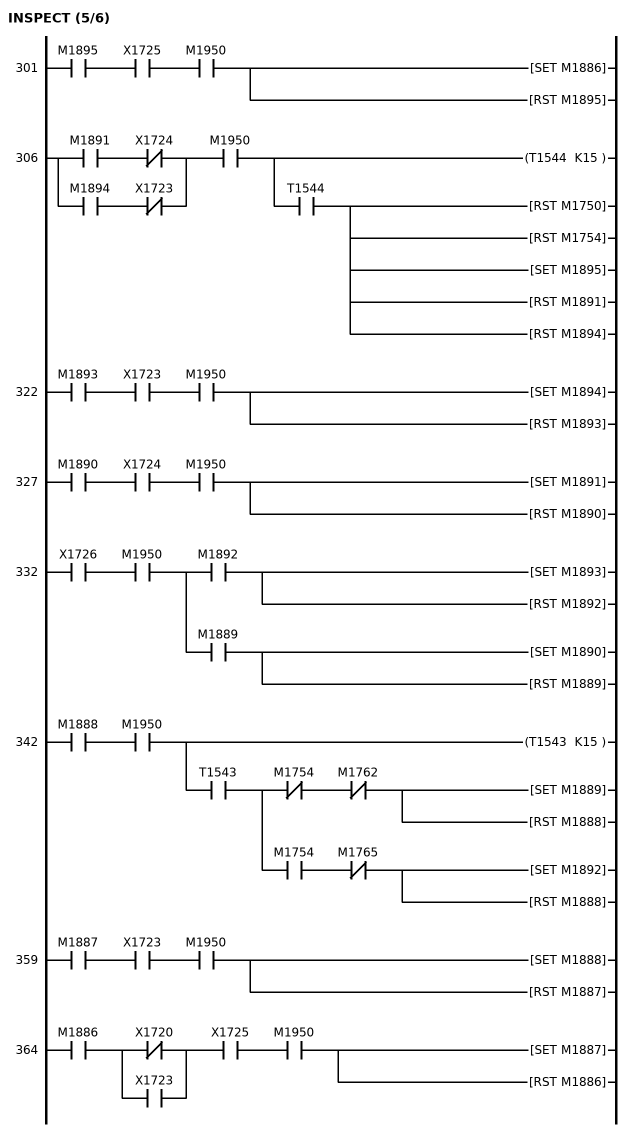
[picture p24: ladder of INSPECT, rungs at steps 301 to 364]
301   LD      M1895
      AND     X1725
      AND     M1950
      SET     M1886
      RST     M1895
306   LD      M1891
      ANI     X1724
      LD      M1894
      ANI     X1723
      ORB
      AND     M1950
      OUT     T1544 K15
      AND     T1544
      RST     M1750
      RST     M1754
      SET     M1895
      RST     M1891
      RST     M1894
322   LD      M1893
      AND     X1723
      AND     M1950
      SET     M1894
      RST     M1893
327   LD      M1890
      AND     X1724
      AND     M1950
      SET     M1891
      RST     M1890
332   LD      X1726
      AND     M1950
      MPS
      AND     M1892
      SET     M1893
      RST     M1892
      MPP
      AND     M1889
      SET     M1890
      RST     M1889
342   LD      M1888
      AND     M1950
      OUT     T1543 K15
      AND     T1543
      MPS
      ANI     M1754
      ANI     M1762
      SET     M1889
      RST     M1888
      MPP
      AND     M1754
      ANI     M1765
      SET     M1892
      RST     M1888
359   LD      M1887
      AND     X1723
      AND     M1950
      SET     M1888
      RST     M1887
364   LD      M1886
      LDI     X1720
      OR      X1723
      ANB
      AND     X1725
      AND     M1950
      SET     M1887
      RST     M1886
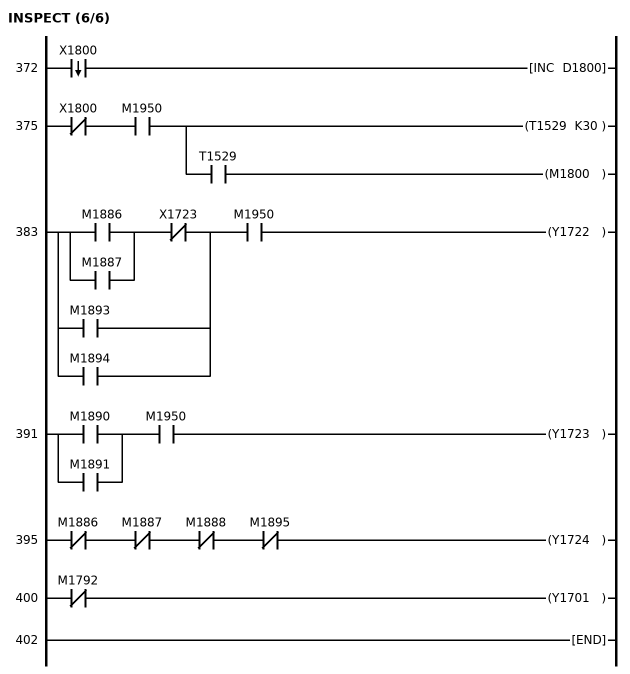
372   LDF     X1800
      INC     D1800
375   LDI     X1800
      AND     M1950
      OUT     T1529 K30
      AND     T1529
      OUT     M1800
383   LD      M1886
      OR      M1887
      ANI     X1723
      LD      M1893
      OR      M1894
      ORB
      AND     M1950
      OUT     Y1722
391   LD      M1890
      OR      M1891
      AND     M1950
      OUT     Y1723
395   LDI     M1886
      ANI     M1887
      ANI     M1888
      ANI     M1895
      OUT     Y1724
400   LDI     M1792
      OUT     Y1701
402   END
END_PROGRAM

PROGRAM RETEST
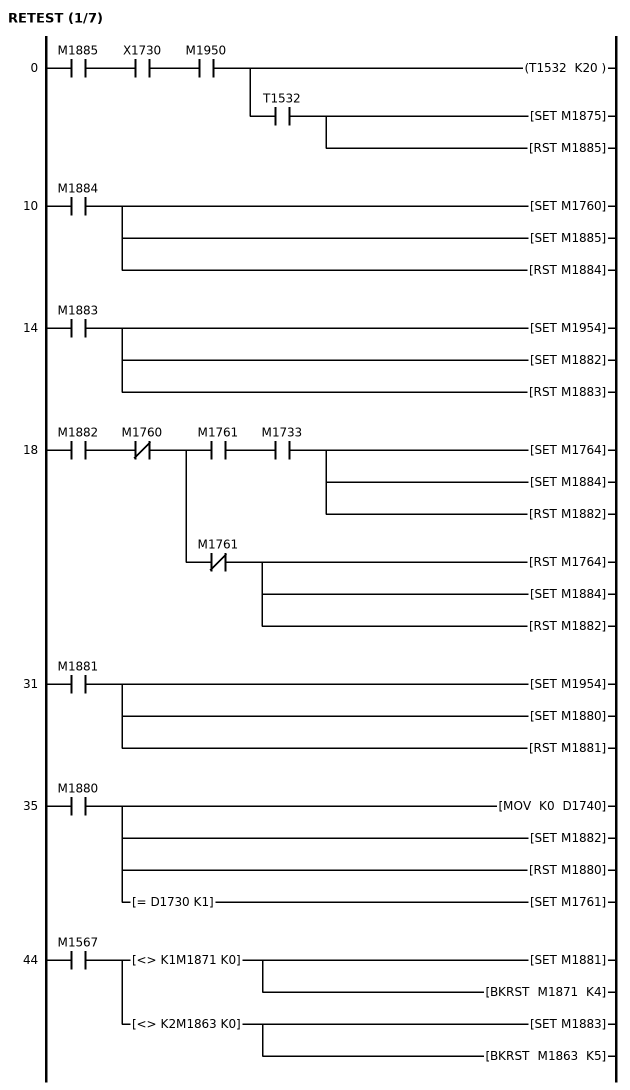
0     LD      M1885
      AND     X1730
      AND     M1950
      OUT     T1532 K20
      AND     T1532
      SET     M1875
      RST     M1885
10    LD      M1884
      SET     M1760
      SET     M1885
      RST     M1884
14    LD      M1883
      SET     M1954
      SET     M1882
      RST     M1883
18    LD      M1882
      ANI     M1760
      MPS
      AND     M1761
      AND     M1733
      SET     M1764
      SET     M1884
      RST     M1882
      MPP
      ANI     M1761
      RST     M1764
      SET     M1884
      RST     M1882
31    LD      M1881
      SET     M1954
      SET     M1880
      RST     M1881
35    LD      M1880
      MOV     K0 D1740
      SET     M1882
      RST     M1880
      AND=    D1730 K1
      SET     M1761
44    LD      M1567
      MPS
      AND<>   K1M1871 K0
      SET     M1881
      BKRST   M1871 K4
      MPP
      AND<>   K2M1863 K0
      SET     M1883
      BKRST   M1863 K5
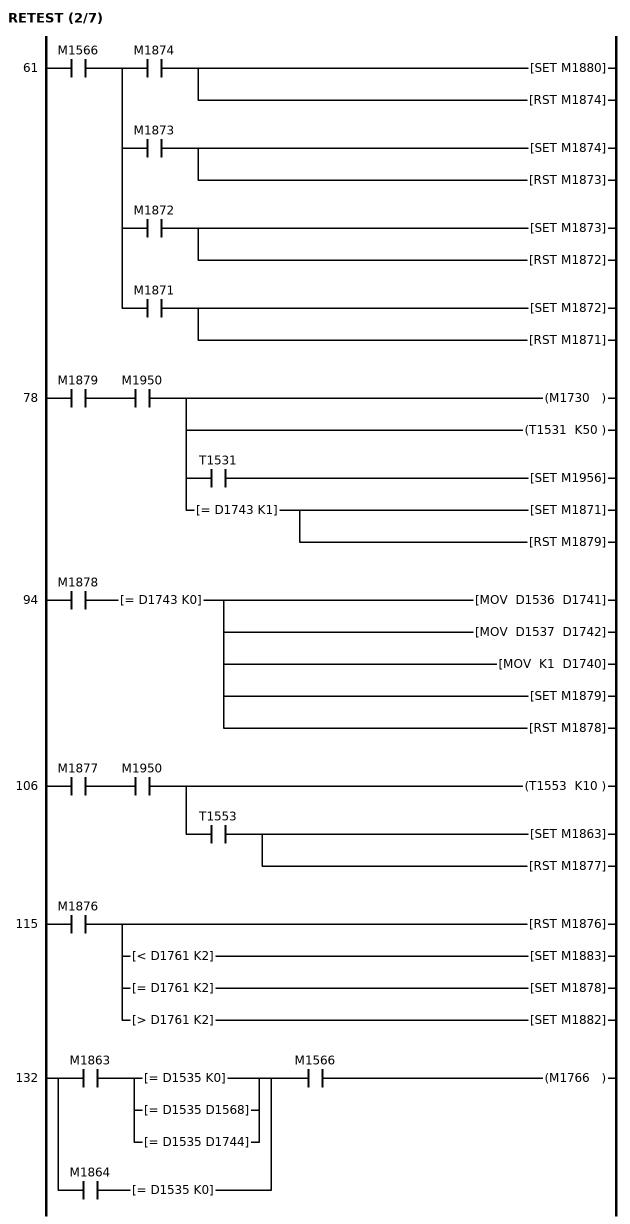
61    LD      M1566
      MPS
      AND     M1874
      SET     M1880
      RST     M1874
      MRD
      AND     M1873
      SET     M1874
      RST     M1873
      MRD
      AND     M1872
      SET     M1873
      RST     M1872
      MPP
      AND     M1871
      SET     M1872
      RST     M1871
78    LD      M1879
      AND     M1950
      OUT     M1730
      OUT     T1531 K50
      MPS
      AND     T1531
      SET     M1956
      MPP
      AND=    D1743 K1
      SET     M1871
      RST     M1879
94    LD      M1878
      AND=    D1743 K0
      MOV     D1536 D1741
      MOV     D1537 D1742
      MOV     K1 D1740
      SET     M1879
      RST     M1878
106   LD      M1877
      AND     M1950
      OUT     T1553 K10
      AND     T1553
      SET     M1863
      RST     M1877
115   LD      M1876
      RST     M1876
      MPS
      AND<    D1761 K2
      SET     M1883
      MRD
      AND=    D1761 K2
      SET     M1878
      MPP
      AND>    D1761 K2
      SET     M1882
132   LD      M1863
      LD=     D1535 K0
      OR=     D1535 D1568
      OR=     D1535 D1744
      ANB
      LD      M1864
      AND=    D1535 K0
      ORB
      AND     M1566
      OUT     M1766
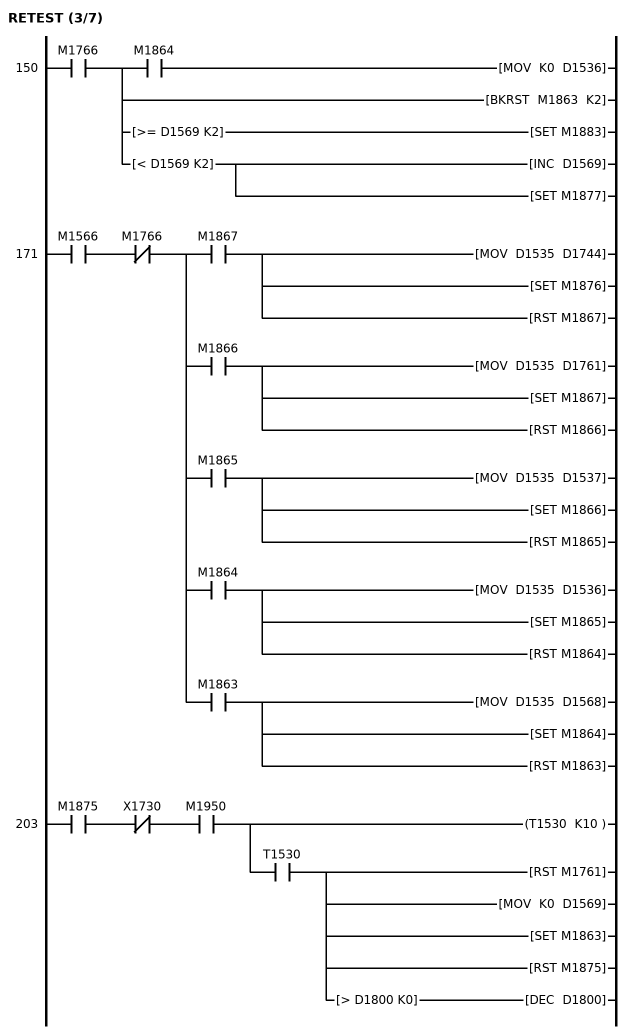
150   LD      M1766
      MPS
      AND     M1864
      MOV     K0 D1536
      MPP
      BKRST   M1863 K2
      MPS
      AND>=   D1569 K2
      SET     M1883
      MPP
      AND<    D1569 K2
      INC     D1569
      SET     M1877
171   LD      M1566
      ANI     M1766
      MPS
      AND     M1867
      MOV     D1535 D1744
      SET     M1876
      RST     M1867
      MRD
      AND     M1866
      MOV     D1535 D1761
      SET     M1867
      RST     M1866
      MRD
      AND     M1865
      MOV     D1535 D1537
      SET     M1866
      RST     M1865
      MRD
      AND     M1864
      MOV     D1535 D1536
      SET     M1865
      RST     M1864
      MPP
      AND     M1863
      MOV     D1535 D1568
      SET     M1864
      RST     M1863
203   LD      M1875
      ANI     X1730
      AND     M1950
      OUT     T1530 K10
      AND     T1530
      RST     M1761
      MOV     K0 D1569
      SET     M1863
      RST     M1875
      AND>    D1800 K0
      DEC     D1800
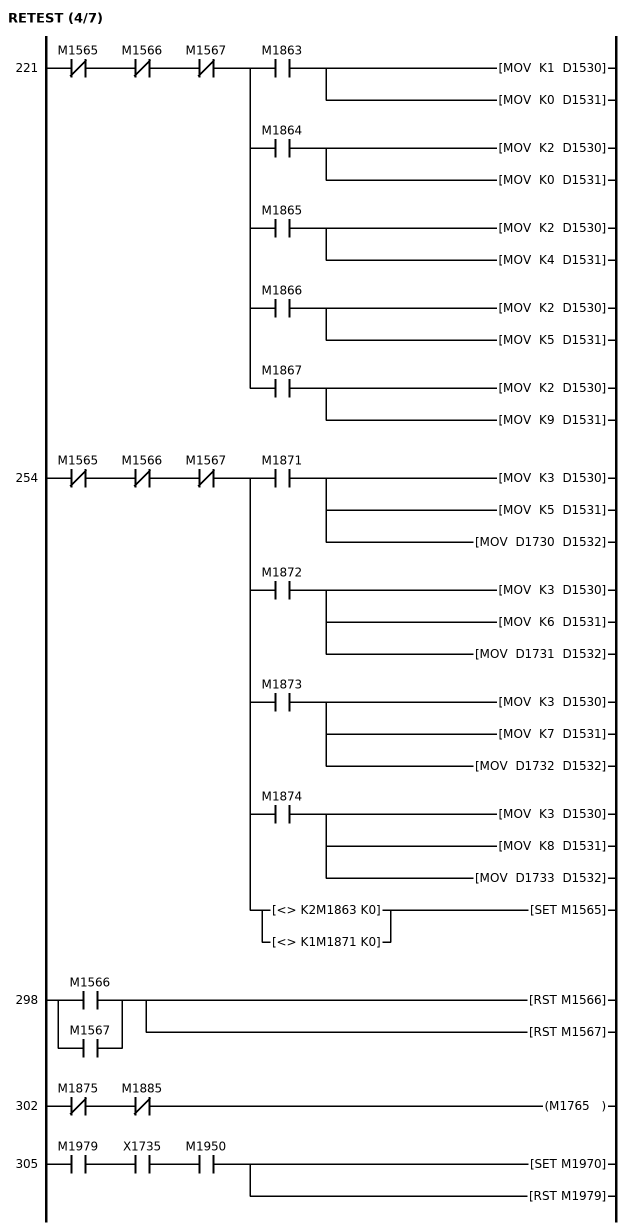
221   LDI     M1565
      ANI     M1566
      ANI     M1567
      MPS
      AND     M1863
      MOV     K1 D1530
      MOV     K0 D1531
      MRD
      AND     M1864
      MOV     K2 D1530
      MOV     K0 D1531
      MRD
      AND     M1865
      MOV     K2 D1530
      MOV     K4 D1531
      MRD
      AND     M1866
      MOV     K2 D1530
      MOV     K5 D1531
      MPP
      AND     M1867
      MOV     K2 D1530
      MOV     K9 D1531
254   LDI     M1565
      ANI     M1566
      ANI     M1567
      MPS
      AND     M1871
      MOV     K3 D1530
      MOV     K5 D1531
      MOV     D1730 D1532
      MRD
      AND     M1872
      MOV     K3 D1530
      MOV     K6 D1531
      MOV     D1731 D1532
      MRD
      AND     M1873
      MOV     K3 D1530
      MOV     K7 D1531
      MOV     D1732 D1532
      MRD
      AND     M1874
      MOV     K3 D1530
      MOV     K8 D1531
      MOV     D1733 D1532
      MPP
      LD<>    K2M1863 K0
      OR<>    K1M1871 K0
      ANB
      SET     M1565
298   LD      M1566
      OR      M1567
      RST     M1566
      RST     M1567
302   LDI     M1875
      ANI     M1885
      OUT     M1765
305   LD      M1979
      AND     X1735
      AND     M1950
      SET     M1970
      RST     M1979
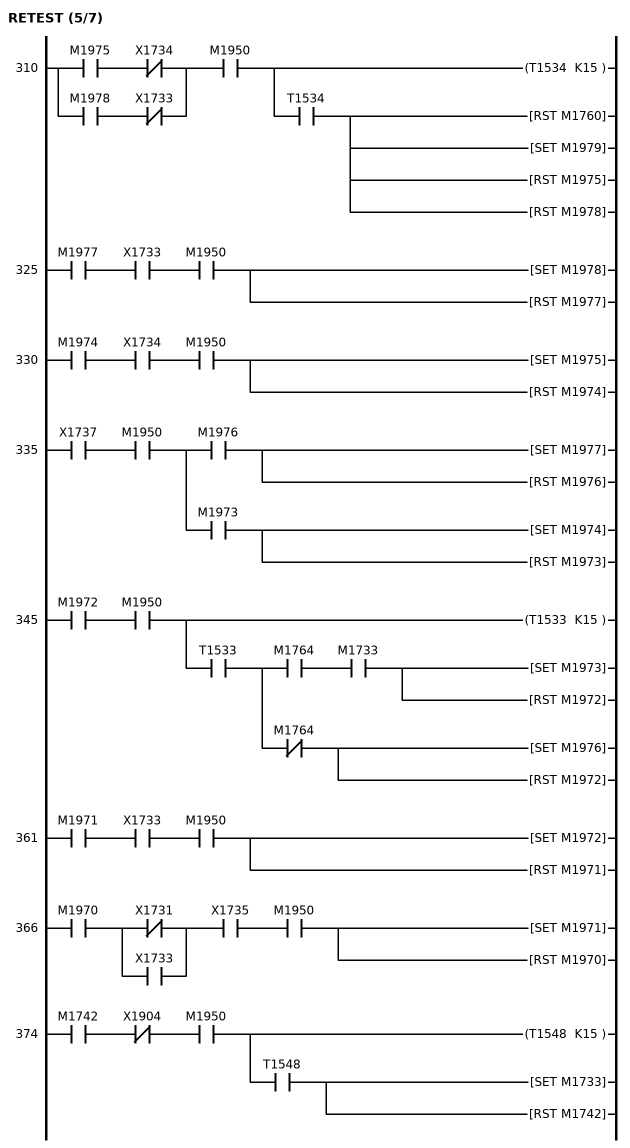
310   LD      M1975
      ANI     X1734
      LD      M1978
      ANI     X1733
      ORB
      AND     M1950
      OUT     T1534 K15
      AND     T1534
      RST     M1760
      SET     M1979
      RST     M1975
      RST     M1978
325   LD      M1977
      AND     X1733
      AND     M1950
      SET     M1978
      RST     M1977
330   LD      M1974
      AND     X1734
      AND     M1950
      SET     M1975
      RST     M1974
335   LD      X1737
      AND     M1950
      MPS
      AND     M1976
      SET     M1977
      RST     M1976
      MPP
      AND     M1973
      SET     M1974
      RST     M1973
345   LD      M1972
      AND     M1950
      OUT     T1533 K15
      AND     T1533
      MPS
      AND     M1764
      AND     M1733
      SET     M1973
      RST     M1972
      MPP
      ANI     M1764
      SET     M1976
      RST     M1972
361   LD      M1971
      AND     X1733
      AND     M1950
      SET     M1972
      RST     M1971
366   LD      M1970
      LDI     X1731
      OR      X1733
      ANB
      AND     X1735
      AND     M1950
      SET     M1971
      RST     M1970
374   LD      M1742
      ANI     X1904
      AND     M1950
      OUT     T1548 K15
      AND     T1548
      SET     M1733
      RST     M1742
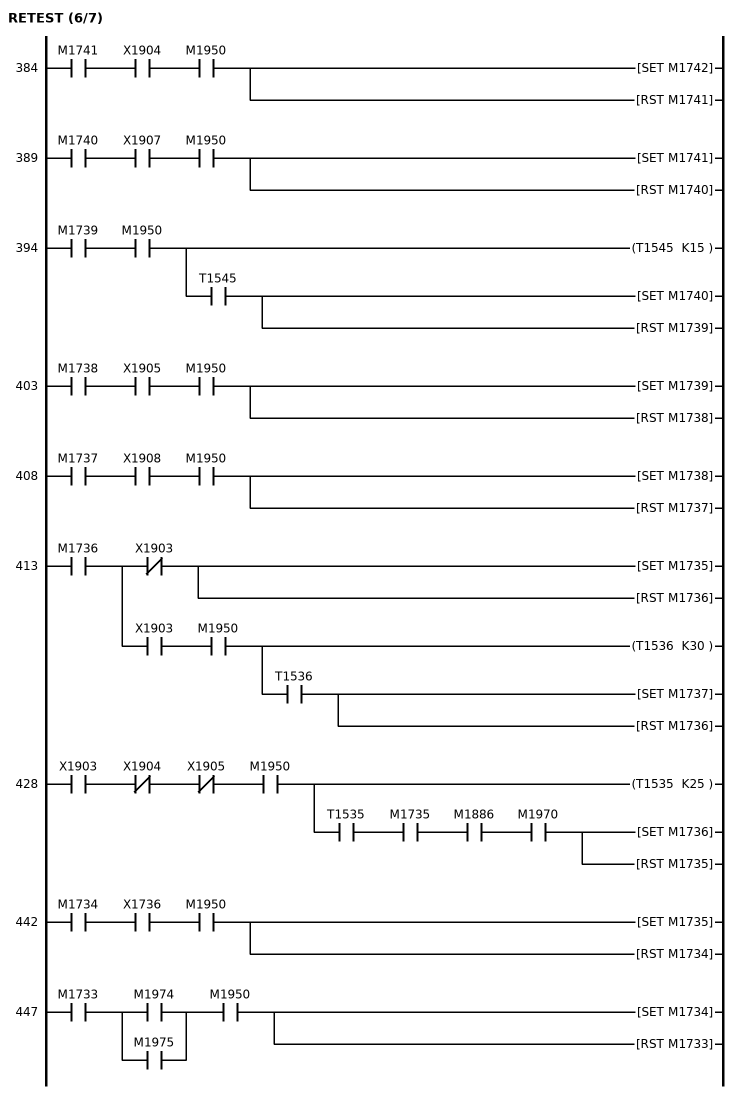
384   LD      M1741
      AND     X1904
      AND     M1950
      SET     M1742
      RST     M1741
389   LD      M1740
      AND     X1907
      AND     M1950
      SET     M1741
      RST     M1740
394   LD      M1739
      AND     M1950
      OUT     T1545 K15
      AND     T1545
      SET     M1740
      RST     M1739
403   LD      M1738
      AND     X1905
      AND     M1950
      SET     M1739
      RST     M1738
408   LD      M1737
      AND     X1908
      AND     M1950
      SET     M1738
      RST     M1737
413   LD      M1736
      MPS
      ANI     X1903
      SET     M1735
      RST     M1736
      MPP
      AND     X1903
      AND     M1950
      OUT     T1536 K30
      AND     T1536
      SET     M1737
      RST     M1736
428   LD      X1903
      ANI     X1904
      ANI     X1905
      AND     M1950
      OUT     T1535 K25
      AND     T1535
      AND     M1735
      AND     M1886
      AND     M1970
      SET     M1736
      RST     M1735
442   LD      M1734
      AND     X1736
      AND     M1950
      SET     M1735
      RST     M1734
447   LD      M1733
      LD      M1974
      OR      M1975
      ANB
      AND     M1950
      SET     M1734
      RST     M1733
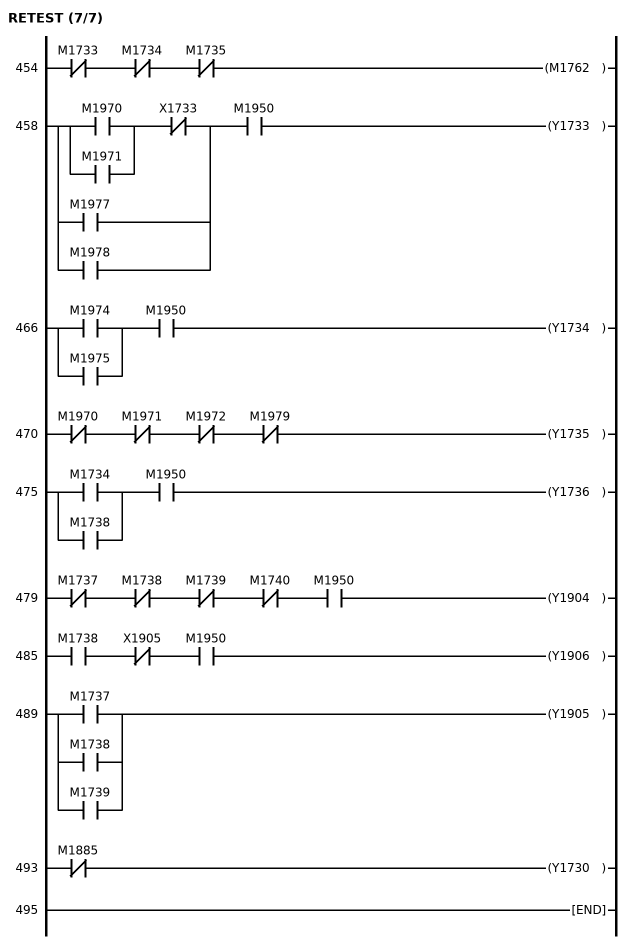
454   LDI     M1733
      ANI     M1734
      ANI     M1735
      OUT     M1762
458   LD      M1970
      OR      M1971
      ANI     X1733
      LD      M1977
      OR      M1978
      ORB
      AND     M1950
      OUT     Y1733
466   LD      M1974
      OR      M1975
      AND     M1950
      OUT     Y1734
470   LDI     M1970
      ANI     M1971
      ANI     M1972
      ANI     M1979
      OUT     Y1735
475   LD      M1734
      OR      M1738
      AND     M1950
      OUT     Y1736
479   LDI     M1737
      ANI     M1738
      ANI     M1739
      ANI     M1740
      AND     M1950
      OUT     Y1904
485   LD      M1738
      ANI     X1905
      AND     M1950
      OUT     Y1906
489   LD      M1737
      OR      M1738
      OR      M1739
      OUT     Y1905
493   LDI     M1885
      OUT     Y1730
495   END
END_PROGRAM

PROGRAM DRIVE
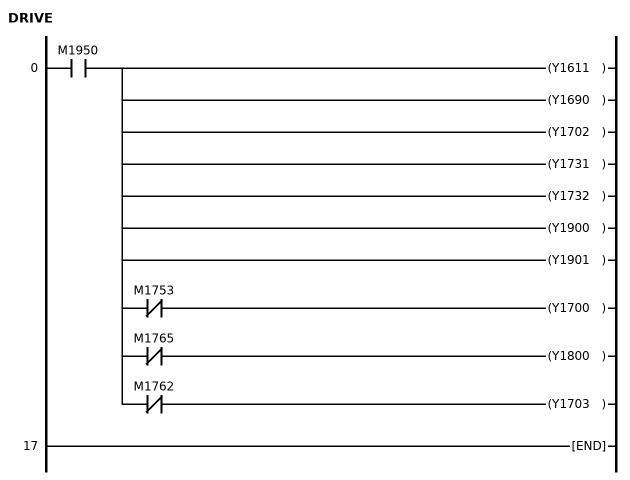
0     LD      M1950
      OUT     Y1611
      OUT     Y1690
      OUT     Y1702
      OUT     Y1731
      OUT     Y1732
      OUT     Y1900
      OUT     Y1901
      MPS
      ANI     M1753
      OUT     Y1700
      MRD
      ANI     M1765
      OUT     Y1800
      MPP
      ANI     M1762
      OUT     Y1703
17    END
END_PROGRAM

PROGRAM COUNTER
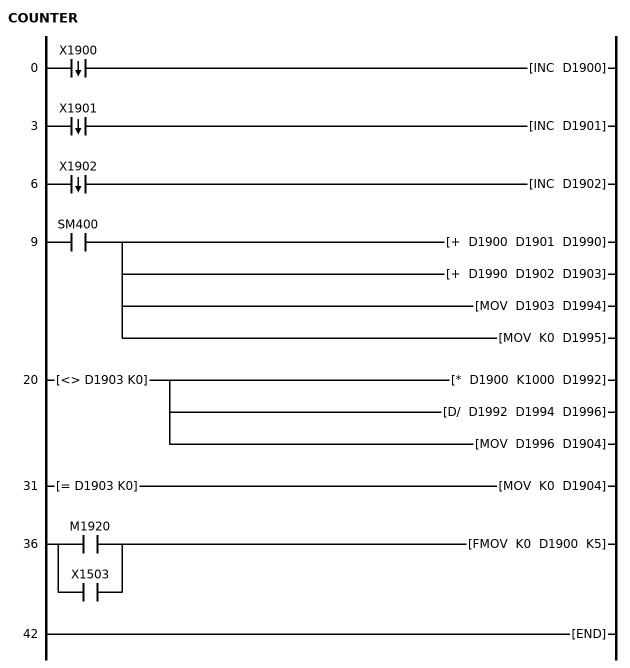
0     LDF     X1900
      INC     D1900
3     LDF     X1901
      INC     D1901
6     LDF     X1902
      INC     D1902
9     LD      SM400
      +       D1900 D1901 D1990
      +       D1990 D1902 D1903
      MOV     D1903 D1994
      MOV     K0 D1995
20    LD<>    D1903 K0
      *       D1900 K1000 D1992
      D/      D1992 D1994 D1996
      MOV     D1996 D1904
31    LD=     D1903 K0
      MOV     K0 D1904
36    LD      M1920
      OR      X1503
      FMOV    K0 D1900 K5
42    END
END_PROGRAM

PROGRAM LAMP
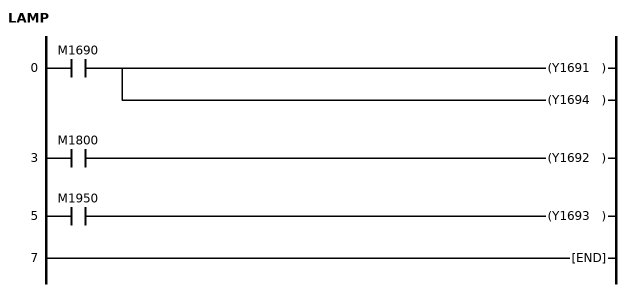
0     LD      M1690
      OUT     Y1691
      OUT     Y1694
3     LD      M1800
      OUT     Y1692
5     LD      M1950
      OUT     Y1693
7     END
END_PROGRAM
